Staubli VAL3: Lab2A_new.dtx


